Fanuc KAREL source: kx00013.KL

-- PROVISIONAL review KL for V770-1; original PC SHA256 19ae525b0b735778486d48a1a95155b37c781fb571f23a4c0c35f15d3b0d16bd
-- Incomplete behavior may be omitted. Consult companion uncertainty JSON. Do not deploy.
PROGRAM KX00013
%NOLOCKGROUP
VAR
  I : INTEGER
  J : INTEGER
  B : BOOLEAN
  F : FILE
  S : STRING[80]
-- UNRESOLVED_DECL P type=000102
BEGIN
  -- UNRESOLVED_PC offsets 5-7; opcodes 9C,4E
  -- UNRESOLVED_PC offsets 12-16; opcodes 7F
END KX00013
